// TIA Portal V21 export
// export: Created 2026-08-21T20:18:49.3042341Z, ExportSetting None, DisplayName Totally Integrated Automation Portal, DisplayVersion V21, DisplayName STEP 7 Professional, DisplayVersion V21, DisplayName STEP 7 Safety, DisplayVersion V21, DisplayName Tech WebApplication, DisplayVersion V21, DisplayName WinCC Basic/Comfort/Advanced, DisplayVersion V21, DisplayName WinCC Professional, DisplayVersion V21, DisplayName WinCC Unified, DisplayVersion V21
FUNCTION_BLOCK "Volumeflow"   // FB1, SCL
{ S7_Optimized_Access := 'TRUE' }
// stored: MemoryReserve 100, SetENOAutomatically false
   VAR_INPUT
      Enable : Bool;
      Release_Spd : Int;
      T_Release : Real;
      Raw_Scale { ExternalAccessible := 'False'; ExternalVisible := 'False'; ExternalWritable := 'False'} : "ScaVal_Raw";
   END_VAR
   VAR_OUTPUT
      Liter : Real;
      Liters_Raw : Int;
   END_VAR
   VAR
      pi : Real := 3.1415;
      r : Real := 0.5;
   END_VAR
   VAR_TEMP
      Release_Spd_Raw : Real;
      Release_Spd_Real : Real;
   END_VAR
   // Raw_Scale.High := 27648;
   // Raw_Scale.Low := 0;
BEGIN
   IF #Enable = FALSE THEN
       #Liter := 0;
       #Liters_Raw := 0;
       RETURN;
   END_IF;
   #Release_Spd_Real := INT_TO_REAL(#Release_Spd);
   #Release_Spd_Raw := (#Release_Spd_Real / 27648) * 100;
   //Volume flow in liter (dm^2 == l)
   #Liter := #T_Release * #Release_Spd_Raw * #pi * #r * #r * 4;
   #Liters_Raw := (#Liter/32) * #Raw_Scale.High;
END_FUNCTION_BLOCK
